Staubli VAL3: hmiClose.pgx

public program hmiClose()
  local bool l_bOut
begin
  delay(0.2)
  utCtn_Message.Appearance.bVisibility=true
  //
  l_bOut=false
  nClock=clock()
  do
    if utCtn_Message.Appearance.bVisibility==true
      if clock()-nClock>=3
        utTxt_popUpMsg.Common.sValue=""
        utCtn_Message.Appearance.bVisibility=false
        l_bOut=true
      endIf
      if utBtn_OK.Events.bClick==true
        utBtn_OK.Events.bClick=false
        utTxt_popUpMsg.Common.sValue=""
        utCtn_Message.Appearance.bVisibility=false
        l_bOut=true
      endIf
    endIf
    delay(0)
  until l_bOut
end
